Fanuc KAREL source: KT00571.KL

PROGRAM KT00571
%NOLOCKGROUP
VAR
  R1: REAL
  V2: VECTOR
  OUT: VECTOR
BEGIN
  R1 = 2.0
    V2.Y = 2.0
  OUT = R1 + V2
END KT00571
